(* PLC project g_pump_alternation, Anonymous Benchmark Suite 1.0 *)
(* stored: creationDateTime 2026-08-28T00:00:00 *)

PROGRAM g_pump_alternation
  VAR_INPUT
    LevelHigh : BOOL;
    LevelLow : BOOL;
  END_VAR
  VAR_OUTPUT
    Call : BOOL;
    Duty : BOOL;
    PumpA : BOOL;
    PumpB : BOOL;
  END_VAR

(* LD diagram, written out as Structured Text *)
Call := (Call OR LevelHigh) AND NOT LevelLow;
Duty := Duty AND NOT LevelLow OR NOT Duty AND LevelLow;
PumpA := Call AND NOT Duty;
PumpB := Call AND Duty;
END_PROGRAM

CONFIGURATION Config0
  RESOURCE Res0 ON PLC
    TASK tcyclic(INTERVAL := T#10ms, PRIORITY := 0);
    PROGRAM inst0 WITH tcyclic : g_pump_alternation;
  END_RESOURCE
END_CONFIGURATION
